// TIA Portal V20 export
VAR_GLOBAL   // PLC tag table "Safety_nicht_F"
   DE_Ueberspannungsschutz_OK AT %I1.0 : Bool;   // DE +SK1-5F1 Überspannungsschutz
   DE_Selektivmodul_OK AT %I1.1 : Bool;   // DE +HS1=AN-22T1 Selektivmodul
   DE_Rueckfuehrung_Tuer_1 AT %I1.2 : Bool;   // DE +Feld=STÜR -921S1 Rückführung Tür 1 ist nicht verriegelt
   DE_Rueckfuehrung_Tuer_2 AT %I1.3 : Bool;   // DE +Feld=STÜR -921S2 Rückführung Tür 2 ist nicht verriegelt (Option)
   DE_Extern_IN1 AT %I1.4 : Bool;   // DE +SK2-911X1 Externe Schnittstelle von Messgerät
   DE_Extern_IN2 AT %I1.5 : Bool;   // DE +SK2-911X1 Externe Schnittstelle von Messgerät
   DE_Extern_IN3 AT %I1.6 : Bool;   // DE +SK2-911X1 Externe Schnittstelle von Messgerät
   "DE_NOT-HALT_Schuetz_Rueckf" AT %I0.0 : Bool;   // DE + HS1=AAS-146K1 NOT-HALT Schütz Rückführung
   "DE_NOT-HALT_Tuere_1_RST_Rueckf" AT %I0.1 : Bool;   // DE + _______NOT-HALT Türe 1 RST Rückführung
   "DE_NOT-HALT_Tuere_1_Rueckf" AT %I0.2 : Bool;   // DE + HS1=AAS-148K1 NOT-HALT Türe 1 Rückführung
   "DE_NOT-HALT_Tuere_2_RST_Rueckf" AT %I0.3 : Bool;   // DE + _______NOT-HALT Türe 2 RST Rückführung
   "DE_NOT-HALT_Tuere_2_Rueckf" AT %I0.4 : Bool;   // DE + _______NOT-HALT Türe 2 Rückführung
   "DE_NOT-HALT_Roboter_Rueckf" AT %I0.5 : Bool;   // DE + _______NOT-HALT Roboter Rückführung
   DE_Sichere_Bewegung_Rueckf AT %I0.6 : Bool;   // DE + _______Sichere Bewegung Rückführung
   DE_Antriebe_Rueckf AT %I0.7 : Bool;   // DE +SK2=ANT-2001T1/-2001T2/2001T3/-2101T1 Antriebe Rückführung
   DE_Extern_IN4 AT %I1.7 : Bool;   // DE +SK2-911X1 Externe Schnittstelle von Messgerät
END_VAR
